// TIA Portal V20 export
Screen "SafetyZone04Overview"  1276x673
  ScreenItem "Button_Overview_LegendᆉY2" at 1185,2 size 90x60  Type=HmiButton
  ScreenItem "Button_Back" at 2,4 size 90x60  Type=HmiButton
  ScreenItem "Line_Header_X0_Y64" at -11,64 size 1280x0  Type=HmiLine
  ScreenItem "Graphic view_15" at 314,334 size 42x35  Type=HmiGraphicView
  ScreenItem "Rectangle_11" at 1176,204 size 148x10  Type=HmiRectangle
  ScreenItem "Rectangle_13" at 27,552 size 468x8  Type=HmiRectangle
  ScreenItem "图形 IO 域_26" at 548,497 size 15x122  Type=HmiSymbolicIOField
  ScreenItem "Button_Overview_LegendᆉY2_1" at 1092,2 size 90x60  Type=HmiButton
  ScreenItem "Button_Overview_LegendᆉY2_2" at 986,2 size 103x60  Type=HmiButton
  ScreenItem "Emerg_3" at 731,83 size 52x56  Type=HmiSymbolicIOField
  ScreenItem "Title_ScreenOverview_X390_Y2_1" at 384,4 size 510x57  Type=HmiTextBox
  ScreenItem "Graphic view_1" at 946,330 size 42x35  Type=HmiGraphicView
  ScreenItem "Emerg_1" at 334,588 size 52x56  Type=HmiSymbolicIOField
  ScreenItem "Button_Overview_LegendᆉY2_3" at 106,2 size 103x60  Type=HmiButton
  ScreenItem "Faceplate container_16" at 742,306 size 152x87  Type=HmiFaceplateContainer
  ScreenItem "Graphic view_2" at 520,76 size 79x51  Type=HmiGraphicView
  ScreenItem "Graphic view_3" at 521,603 size 79x51  Type=HmiGraphicView
  ScreenItem "Rectangle_1" at 619,552 size 625x9  Type=HmiRectangle
  ScreenItem "图形 IO 域_1" at 553,78 size 15x122  Type=HmiSymbolicIOField
  ScreenItem "Rectangle_2" at 633,137 size 620x9  Type=HmiRectangle
  ScreenItem "Rectangle_3" at 32,135 size 466x9  Type=HmiRectangle
  ScreenItem "符号 IO 域_4" at 355,86 size 43x40  Type=HmiSymbolicIOField
  ScreenItem "Text_15" at 238,83 size 160x40  Type=HmiText
  ScreenItem "符号 IO 域_1" at 991,600 size 43x40  Type=HmiSymbolicIOField
  ScreenItem "Text_1" at 874,597 size 160x40  Type=HmiText
  ScreenItem "Faceplate container_1" at 355,286 size 362x136  Type=HmiFaceplateContainer
  ScreenItem "图形 IO 域_15" at 1244,283 size 15x122  Type=HmiSymbolicIOField
  ScreenItem "Rectangle_5" at 1176,481 size 148x10  Type=HmiRectangle
  ScreenItem "Rectangle_4" at -37,204 size 148x10  Type=HmiRectangle
  ScreenItem "图形 IO 域_2" at 31,283 size 15x122  Type=HmiSymbolicIOField
  ScreenItem "Rectangle_6" at -38,481 size 148x10  Type=HmiRectangle
